Fanuc KAREL source: KA00211.KL

PROGRAM KA00211
%NOLOCKGROUP
VAR
  SRC: ARRAY[4] OF XYZWPR
  DST: ARRAY[4] OF STRING[20]
BEGIN
  DST = SRC
END KA00211
